(* IEC 61131-3 sources: Test-Git_ESME26/TestProgettoESME_26.fbsproj/PacDriveLib Migration/Motion/Positioning/PDL_FB_VarioPosJerk.fb.st^, 6 files *)

(* ---- etPosModeToString.meth.st ---- *)
METHOD PRIVATE etPosModeToString : STRING[10]
VAR_INPUT
	i_etPosMode		: PDL_ET_PosMode;
END_VAR

CASE i_etPosMode OF
	PDL_ET_PosMode.Absolute:
		etPosModeToString := 'Absolute';

	PDL_ET_PosMode.Endless:
		etPosModeToString := 'Endless';

	PDL_ET_PosMode.Relative:
		etPosModeToString := 'Relative';

ELSE
	etPosModeToString := 'Unknown';
END_CASE

(* ---- Init.meth.st ---- *)
{attribute 'hide'}
METHOD PRIVATE Init : BOOL
VAR_INPUT
END_VAR

Init := FALSE;

IF i_ifDrive = 0 THEN
	SetDiagOutput(	i_etDiag	:= GD.ET_Diag.InputParameterInvalid,
					i_etDiagExt := PDL_ET_DiagExt.DriveInvalid,
					i_sMsg		:= 'i_ifDrive - Invalid Interface');
	RETURN;
ELSE
	//get IF_DriveConfig
	xSuccess := __QUERYINTERFACE(i_ifDrive, ifGetParentDevice);
	IF xSuccess AND ifGetParentDevice <> 0 THEN
		ifDeviceAccess := ifGetParentDevice.GetParentDevice();
		xSuccess := __QUERYINTERFACE( ifDeviceAccess, ifDriveConfigAccess );
		IF xSuccess AND ifDriveConfigAccess <> 0 THEN
			ifDriveConfig := ifDriveConfigAccess.DriveConfig;
		END_IF
	END_IF

	xSuccess := __QUERYINTERFACE(ifDeviceAccess, ifDeviceTreeObjectAccess);
	IF xSuccess THEN
		sDriveName := ifDeviceTreeObjectAccess.DeviceTreeObject.Name;
	ELSE
		sDriveName := 'Axis';
	END_IF

	fbHalt.Axis := i_ifDrive;
	fbStop.Axis := i_ifDrive;
	fbMoveAbsolute.Axis := i_ifDrive;
	fbMoveRelative.Axis := i_ifDrive;

END_IF

//i_ifDrive.lrModuloPeriod

Init := TRUE;

(* ---- InputParameterCheck.meth.st ---- *)
METHOD PRIVATE InputParameterCheck : BOOL
VAR_INPUT
END_VAR
VAR
	lrMaxAcc	: LREAL := 0;
	lrMaxVel	: LREAL := 0;
END_VAR

InputParameterCheck := FALSE;

//if IF_DriveConfig is not available -> limits are NOT checked
IF ifDriveConfig <> 0 THEN
	lrMaxAcc := ifDriveConfig.MaxAcc;
	lrMaxVel := ifDriveConfig.MaxVel;
END_IF

IF i_lrVel <= 0  OR (i_lrVel > lrMaxVel AND lrMaxVel <> 0) THEN
		SetDiagOutput(	i_etDiag	:= GD.ET_Diag.InputParameterInvalid,
						i_etDiagExt := PDL_ET_DiagExt.VelRange,
						i_sMsg		:= SE_CTBX.FC_MultiConcat(	i_sString1 := '0 < i_lrVel <= ',
																i_sString2 := TO_STRING( lrMaxVel),
																i_sString3 := '',
																i_sString4 := ''));

ELSIF i_lrAcc <= 0 OR (i_lrAcc > lrMaxAcc AND lrMaxAcc <> 0) THEN
		SetDiagOutput(	i_etDiag	:= GD.ET_Diag.InputParameterInvalid,
						i_etDiagExt := PDL_ET_DiagExt.AccRange,
						i_sMsg		:= SE_CTBX.FC_MultiConcat(	i_sString1 := '0.0 < ',
																i_sString2 := 'i_lrAcc',
																i_sString3 := ' <= ',
																i_sString4 := TO_STRING(lrMaxAcc)
																));

ELSIF i_lrDec <= 0 OR (i_lrDec > lrMaxAcc AND lrMaxAcc <> 0) THEN
		SetDiagOutput(	i_etDiag	:= GD.ET_Diag.InputParameterInvalid,
						i_etDiagExt := PDL_ET_DiagExt.DecRange,
						i_sMsg		:= SE_CTBX.FC_MultiConcat(	i_sString1 := '0.0 < ',
																i_sString2 := 'i_lrDec',
																i_sString3 := ' <= ',
																i_sString4 := TO_STRING(lrMaxAcc)
																));

ELSIF    (i_etPosMode <> PDL_ET_PosMode.Absolute)
	AND  (i_etPosMode <> PDL_ET_PosMode.Relative)
	AND  (i_etPosMode <> PDL_ET_PosMode.Endless)
THEN
	SetDiagOutput(	i_etDiag	:= GD.ET_Diag.InputParameterInvalid,
					i_etDiagExt := PDL_ET_DiagExt.PosModeRange,
					i_sMsg		:= '');

ELSIF i_lrJerk <= 0.0  THEN
	SetDiagOutput(	i_etDiag	:= GD.ET_Diag.InputParameterInvalid,
					i_etDiagExt := PDL_ET_DiagExt.JerkRange,
					i_sMsg		:= '0.0 < i_lrJerk ');
ELSE
	InputParameterCheck := TRUE;
END_IF

//Target-Prüfung fehlt noch

(* ---- RegisterLoggerPoint.meth.st ---- *)
METHOD PUBLIC RegisterLoggerPoint
VAR_INPUT
	i_ifParent		: APL.IF_LoggerPoint;
	i_sName			: STRING[80];
END_VAR
VAR_OUTPUT
	q_etDiag		: GD.ET_Diag := GD.ET_Diag.Ok;
	q_etDiagExt		: PDL_ET_DiagExt := PDL_ET_DiagExt.Ok;
END_VAR
VAR
	etDiagBuffer		: GD.ET_Diag;
	etDiagExtBufferAPL	: APL.ET_DiagExt;
END_VAR

fbLoggerPoint.RegisterLoggerPoint(	i_ifParent		:= i_ifParent,
									i_sName			:= i_sName,
									i_sType			:= 'FB_VarioPosJerk',
									i_sSource		:= 'PDL',
									q_etDiag		=> etDiagBuffer,
									q_etDiagExt		=> etDiagExtBufferAPL);
IF (etDiagBuffer <> GD.ET_Diag.Ok) THEN
	CASE etDiagExtBufferAPL OF
		APL.ET_DiagExt.ParentInvalid:
			q_etDiag := GD.ET_Diag.InputParameterInvalid;
			q_etDiagExt := PDL_ET_DiagExt.ParentInvalid;

		APL.ET_DiagExt.ParentNotRegistered:
			q_etDiag := GD.ET_Diag.InputParameterInvalid;
			q_etDiagExt := PDL_ET_DiagExt.ParentNotRegistered;

		APL.ET_DiagExt.MaxNumberOfLoggerPointsExeeded:
			q_etDiag := GD.ET_Diag.InputParameterInvalid;
			q_etDiagExt := PDL_ET_DiagExt.MaxNumberOfLoggerPointsExeeded;

	ELSE
		q_etDiag := GD.ET_Diag.UnexpectedProgramBehavior;
		q_etdiagExt := PDL_ET_DiagExt.UnexpectedDiagExt;
	END_CASE
END_IF

(* ---- SetDiagOutput.meth.st ---- *)
METHOD PRIVATE SetDiagOutput : BOOL
VAR_INPUT
	i_etDiag	: GD.ET_Diag;
	i_etDiagExt	: PDL_ET_DiagExt;
	i_sMsg		: STRING[80];
END_VAR
VAR
END_VAR

IF i_etDiag <> GD.ET_Diag.Ok THEN
	q_xReady := FALSE;
END_IF
IF q_etDiag = GD.ET_Diag.OK OR i_etDiagExt = PDL_ET_DiagExt.Disabled THEN
	q_etDiag := i_etDiag;
	q_etDiagExt := i_etDiagExt;
	q_sMsg := i_sMsg;

	IF(i_etDiag = GD.ET_Diag.Ok) AND (fbLoggerPoint.etLogLevel >= APL.ET_LogLevel.StatusMessage) THEN
		fbLoggerPoint.AddLogEntry(	i_etLogLevel	:= APL.ET_LogLevel.StatusMessage,
									i_etDiag		:= q_etDiag,
									i_udiDiagExt	:= q_etDiagExt,
									i_sMessage		:= SE_CTBX.FC_MultiConcat(	i_sString1	:= Standard.CONCAT('ET_Diag: ', GD.FC_EtDiagToString(q_etDiag)),
																				i_sString2	:= Standard.CONCAT(' ET_DiagExt: ', PDL_FC_EtDiagExtToString(q_etDiagExt)),
																				i_sString3	:= Standard.CONCAT(' sMsg: ', q_sMsg),
																				i_sString4	:= '')
											);
	ELSIF(i_etDiag = GD.ET_Diag.UnexpectedProgramBehavior) AND (fbLoggerPoint.etLogLevel >= APL.ET_LogLevel.CriticalException) THEN
		fbLoggerPoint.AddLogEntry(	i_etLogLevel	:= APL.ET_LogLevel.CriticalException,
									i_etDiag		:= q_etDiag,
									i_udiDiagExt	:= q_etDiagExt,
									i_sMessage		:= SE_CTBX.FC_MultiConcat(	i_sString1	:= Standard.CONCAT('ET_Diag: ', GD.FC_EtDiagToString(q_etDiag)),
																				i_sString2	:= Standard.CONCAT(' ET_DiagExt: ', PDL_FC_EtDiagExtToString(q_etDiagExt)),
																				i_sString3	:= Standard.CONCAT(' sMsg: ', q_sMsg),
																				i_sString4	:= '')
											);
	ELSIF(i_etDiag <> GD.ET_Diag.Ok) AND (fbLoggerPoint.etLogLevel >= APL.ET_LogLevel.Exception) THEN
		fbLoggerPoint.AddLogEntry(	i_etLogLevel	:= APL.ET_LogLevel.Exception,
									i_etDiag		:= q_etDiag,
									i_udiDiagExt	:= q_etDiagExt,
									i_sMessage		:= SE_CTBX.FC_MultiConcat(	i_sString1	:= Standard.CONCAT('ET_Diag: ', GD.FC_EtDiagToString(q_etDiag)),
																				i_sString2	:= Standard.CONCAT(' ET_DiagExt: ', PDL_FC_EtDiagExtToString(q_etDiagExt)),
																				i_sString3	:= Standard.CONCAT(' sMsg: ', q_sMsg),
																				i_sString4	:= '')
									);
	END_IF
END_IF

(* ---- SetPos.meth.st ---- *)
METHOD PRIVATE SetPos : BOOL
VAR_INPUT
END_VAR

IF i_etPosMode = PDL_ET_PosMode.Endless THEN

	fbSetPos( 	Axis		:= i_ifDrive,
				Execute		:= FALSE);

	fbSetPos( 	Axis		:= i_ifDrive,
				Execute		:= TRUE,
				Position 	:= 0,
				Relative  	:= FALSE
				);

	IF   fbSetPos.Error
	  OR NOT fbSetPos.Done
	THEN
		SetDiagOutput(	i_etDiag	:= GD.ET_Diag.UnexpectedProgramBehavior,
						i_etDiagExt := PDL_ET_DiagExt.UnexpectedFeedback,
						i_sMsg		:= CONCAT('MC_SetPosition.ErrorID: ', TO_STRING(fbSetPos.ErrorID) ));

		fbSetPos( 	Axis		:= i_ifDrive,
					Execute		:= FALSE);
		diState := 0;
		RETURN;
	END_IF

END_IF
